PROGRAM main
  VAR
    SCADA_CALL_FLOOR_1 AT %QX0.0 : BOOL;
    SCADA_CALL_FLOOR_2 AT %QX0.1 : BOOL;
    SCADA_CALL_FLOOR_3 AT %QX0.2 : BOOL;
    SCADA_ELEVATOR_DISABLE AT %QX0.3 : BOOL;
    PUB_ELEVATOR_MOVING AT %QX0.4 : BOOL;
    PUB_ELEVATOR_FAULT AT %QX0.5 : BOOL;
    PUB_CURRENT_FLOOR AT %QW0 : UINT;
    PUB_HEARTBEAT AT %QW1 : UINT;
    PUB_RECONNECT_COUNT AT %QW2 : UINT;
    CALL_FLOOR_1 AT %QX100.0 : BOOL;
    CALL_FLOOR_2 AT %QX100.1 : BOOL;
    CALL_FLOOR_3 AT %QX100.2 : BOOL;
    ELEVATOR_DISABLE AT %QX100.3 : BOOL;
    ELEVATOR_MOVING AT %IX100.0 : BOOL;
    ELEVATOR_FAULT AT %IX100.1 : BOOL;
    CURRENT_FLOOR AT %IW100 : UINT;
    HEARTBEAT AT %IW101 : UINT;
    RECONNECT_COUNT AT %IW102 : UINT;
    CALL_PULSE_TIME : TIME := T#300ms;
    TP0 : TP;
    TP1 : TP;
    TP2 : TP;
  END_VAR

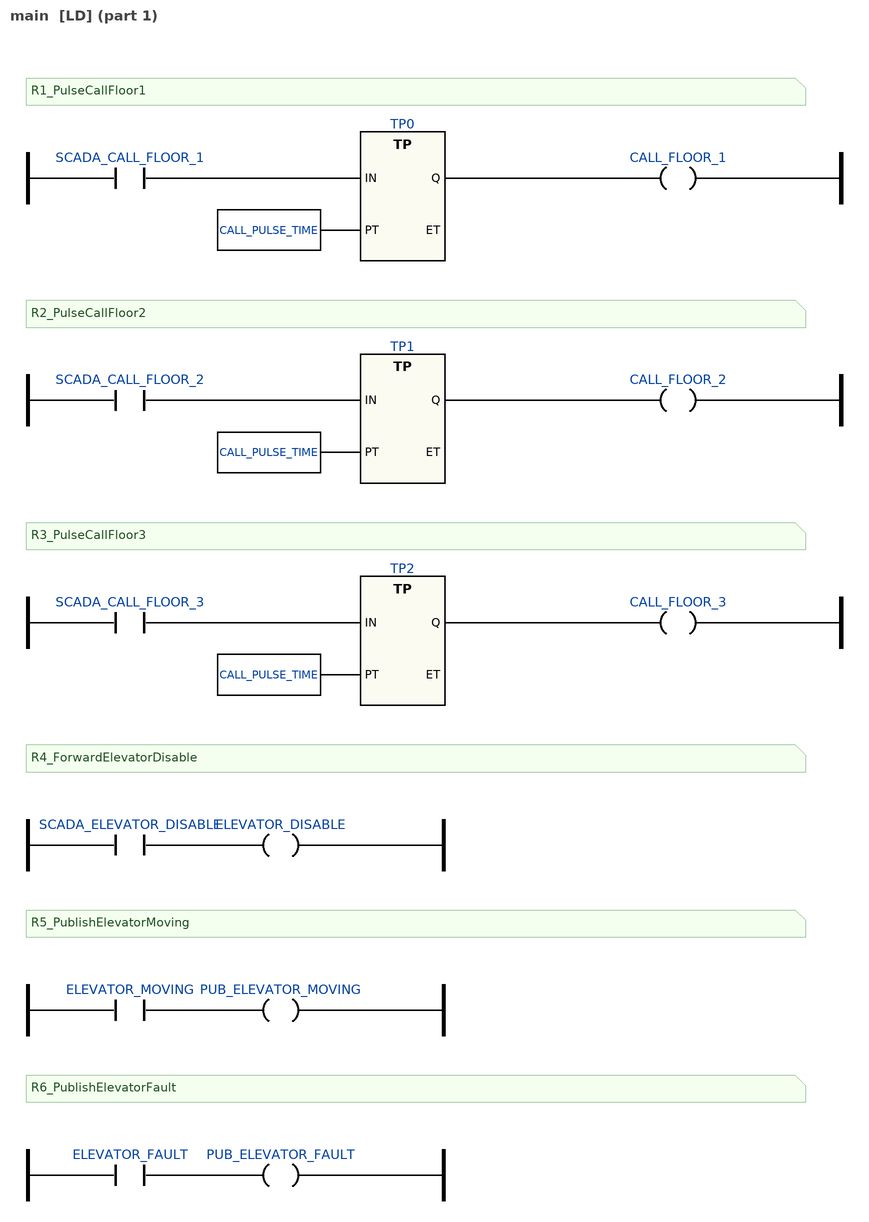
(* LD diagram, written out as Structured Text *)
(* R1_PulseCallFloor1 *)
TP0(IN := SCADA_CALL_FLOOR_1, PT := CALL_PULSE_TIME);
CALL_FLOOR_1 := TP0.Q;
(* R2_PulseCallFloor2 *)
TP1(IN := SCADA_CALL_FLOOR_2, PT := CALL_PULSE_TIME);
CALL_FLOOR_2 := TP1.Q;
(* R3_PulseCallFloor3 *)
TP2(IN := SCADA_CALL_FLOOR_3, PT := CALL_PULSE_TIME);
CALL_FLOOR_3 := TP2.Q;
(* R4_ForwardElevatorDisable *)
ELEVATOR_DISABLE := SCADA_ELEVATOR_DISABLE;
(* R5_PublishElevatorMoving *)
PUB_ELEVATOR_MOVING := ELEVATOR_MOVING;
(* R6_PublishElevatorFault *)
PUB_ELEVATOR_FAULT := ELEVATOR_FAULT;
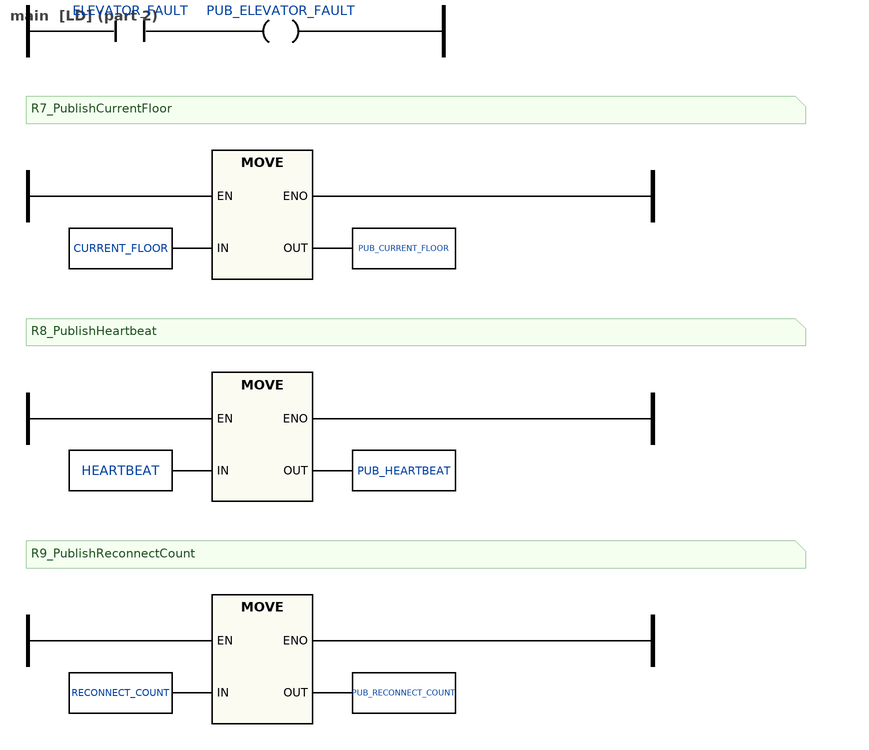
(* R7_PublishCurrentFloor *)
PUB_CURRENT_FLOOR := CURRENT_FLOOR;
(* R8_PublishHeartbeat *)
PUB_HEARTBEAT := HEARTBEAT;
(* R9_PublishReconnectCount *)
PUB_RECONNECT_COUNT := RECONNECT_COUNT;
END_PROGRAM
